Fanuc KAREL source: ko00095.KL

PROGRAM KO00095
%STACKSIZE=65535
%PRIORITY=65535
%NOLOCKGROUP
VAR
P1 : JOINTPOS9
P2 : JOINTPOS9
F : BOOLEAN
OUT : XYZWPREXT
BEGIN
F=TRUE
-- UNSAFE_SOURCE_IR line 11: OUT = MIRROR(convert_jointpos9_to_xyzwprext(P1), convert_jointpos9_to_position(P2), F)
END KO00095
